PROGRAM main
  VAR
    stop : BOOL;
    start : BOOL;
    machine_run : BOOL;
    TOF0 : TOF;
    fan : BOOL;
    high_temp : BOOL;
  END_VAR

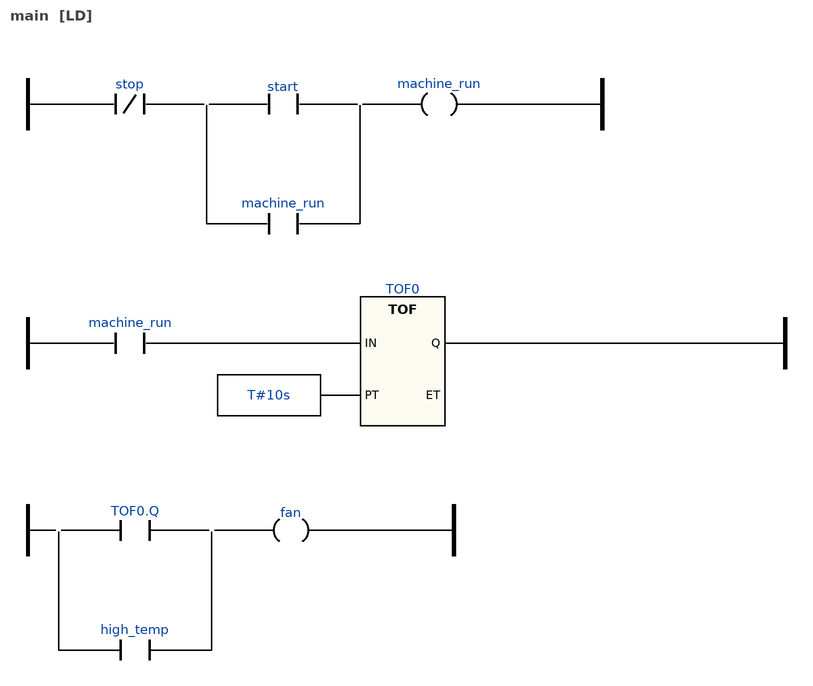
(* LD diagram, written out as Structured Text *)
machine_run := NOT stop AND (start OR machine_run);
fan := TOF0.Q OR high_temp;
TOF0(IN := machine_run, PT := T#10s);
END_PROGRAM
